// TIA Portal project "TrafficLight" (V19)

(* hardware
DEVICE "S7-1200 station_1"  S7-1200 Station
   slot 0: "Rack_0"  S7-1200 Rack  Rack  V1.0
   slot 1: "PLC_1"  CPU 1215C DC/DC/DC  6ES7 215-1AG40-0XB0  V4.6
*)

// ===== PLC "PLC_1"  CPU 1215C DC/DC/DC =====

VAR_GLOBAL   // PLC tag table "Default tag table"
   "emergencyButton" AT %I0.0 : Bool;
   "pedButtonDirB" AT %I0.1 : Bool;
   "pedButtonDirA" AT %I0.2 : Bool;
   "greenDirA" AT %Q0.0 : Bool;
   "yellowDirA" AT %Q0.1 : Bool;
   "redDirA" AT %Q0.2 : Bool;
   "pedGreenDirB" AT %Q0.3 : Bool;
   "pedRedDirB" AT %Q0.4 : Bool;
   "greenDirB" AT %Q0.5 : Bool;
   "yellowDirB" AT %Q0.6 : Bool;
   "redDirB" AT %Q0.7 : Bool;
   "pedGreenDirA" AT %Q1.0 : Bool;
   "pedRedDirA" AT %Q1.1 : Bool;
   "pedReqA" AT %M0.4 : Bool;
   "pedReqB" AT %M0.5 : Bool;
   "emergencyMode" AT %M0.6 : Bool;
   "current_dir" AT %M0.7 : Bool;
   "init_done" AT %M1.0 : Bool;
   "_debug" AT %M1.1 : Bool;
END_VAR

// folder: System blocks/Program resources

DATA_BLOCK "TP_Yellow_Phase_1"   // DB2
{ S7_Optimized_Access := 'TRUE' }
AUTHOR : Simatic
FAMILY : IEC
NAME : IEC_TMR
VERSION : 1.0
// stored: InstanceOfName IEC_TIMER
"IEC_TIMER"
BEGIN
END_DATA_BLOCK

DATA_BLOCK "TP_Yellow_Phase_2"   // DB3
{ S7_Optimized_Access := 'TRUE' }
AUTHOR : Simatic
FAMILY : IEC
NAME : IEC_TMR
VERSION : 1.0
// stored: InstanceOfName IEC_TIMER
"IEC_TIMER"
BEGIN
END_DATA_BLOCK

DATA_BLOCK "tp_main_loop"   // DB6
{ S7_Optimized_Access := 'TRUE' }
AUTHOR : Simatic
FAMILY : IEC
NAME : IEC_TMR
VERSION : 1.0
// stored: InstanceOfName IEC_TIMER
"IEC_TIMER"
BEGIN
END_DATA_BLOCK

DATA_BLOCK "ton_main_loop"   // DB7
{ S7_Optimized_Access := 'TRUE' }
AUTHOR : Simatic
FAMILY : IEC
NAME : IEC_TMR
VERSION : 1.0
// stored: InstanceOfName IEC_TIMER
"IEC_TIMER"
BEGIN
END_DATA_BLOCK

DATA_BLOCK "tp_main_loop_2"   // DB8
{ S7_Optimized_Access := 'TRUE' }
AUTHOR : Simatic
FAMILY : IEC
NAME : IEC_TMR
VERSION : 1.0
// stored: InstanceOfName IEC_TIMER
"IEC_TIMER"
BEGIN
END_DATA_BLOCK

// folder: (top level)

FUNCTION "ped_request" : Void   // FC1, LAD
{ S7_Optimized_Access := 'TRUE' }
VERSION : 0.1
   VAR_INPUT
      pred_A_or_B : String;
      ped_button : Bool;
      ped_req : Bool;
      ped_green : Bool;
      ped_red : Bool;
      dir_red : Bool;
   END_VAR
   VAR_OUTPUT
      o_ped_red : Bool;
      o_ped_green : Bool;
      o_ped_req : Bool;
   END_VAR
   VAR_TEMP
      r_trig_Q : Bool;
   END_VAR
   VAR_TEMP   // added for the SCL form of the ladder/FBD networks
      _w1 : Bool;
   END_VAR
BEGIN

REGION Network 1
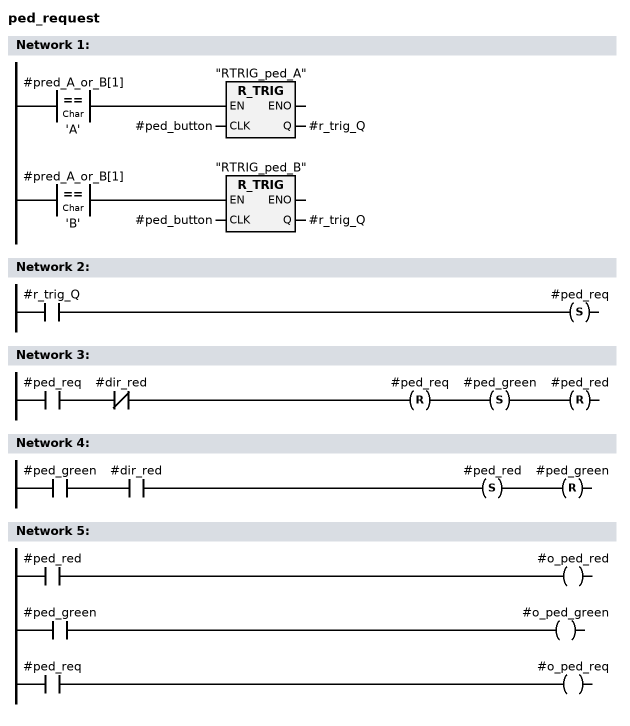
   IF #pred_A_or_B[1] = 'A' THEN
       "RTRIG_ped_A"(CLK := #ped_button, Q => #r_trig_Q);   // R_TRIG
   END_IF;
   IF #pred_A_or_B[1] = 'B' THEN
       "RTRIG_ped_B"(CLK := #ped_button, Q => #r_trig_Q);   // R_TRIG
   END_IF;
END_REGION

REGION Network 2
   RUNG wire#powerrail
      Contact( #r_trig_Q )
      S_Coil( #ped_req )
   END_RUNG
   // the same network as SCL:
   IF #r_trig_Q THEN #ped_req := TRUE; END_IF;
END_REGION

REGION Network 3
   RUNG wire#powerrail
      Contact( #ped_req )
      I_Contact( #dir_red )
      R_Coil( #ped_req )
      S_Coil( #ped_green )
      R_Coil( #ped_red )
   END_RUNG
   // the same network as SCL:
   #_w1 := #ped_req AND NOT #dir_red;
   IF #_w1 THEN
       #ped_req := FALSE;
       #ped_green := TRUE;
       #ped_red := FALSE;
   END_IF;
END_REGION

REGION Network 4
   RUNG wire#powerrail
      Contact( #ped_green )
      Contact( #dir_red )
      S_Coil( #ped_red )
      R_Coil( #ped_green )
   END_RUNG
   // the same network as SCL:
   IF #ped_green AND #dir_red THEN
       #ped_red := TRUE;
       #ped_green := FALSE;
   END_IF;
END_REGION

REGION Network 5
   RUNG wire#powerrail
      Contact( #ped_red )
      Coil( #o_ped_red )
   END_RUNG
   RUNG wire#powerrail
      Contact( #ped_green )
      Coil( #o_ped_green )
   END_RUNG
   RUNG wire#powerrail
      Contact( #ped_req )
      Coil( #o_ped_req )
   END_RUNG
   // the same network as SCL:
   #o_ped_red := #ped_red;
   #o_ped_green := #ped_green;
   #o_ped_req := #ped_req;
END_REGION
END_FUNCTION

FUNCTION "emerg" : Void   // FC2, LAD
{ S7_Optimized_Access := 'TRUE' }
VERSION : 0.1
   VAR_TEMP
      null_p : Bool;
   END_VAR
   VAR_TEMP   // added for the SCL form of the ladder/FBD networks
      _w1 : Bool;
      _w2 : Bool;
   END_VAR
BEGIN

REGION Network 1
   // Notice button click
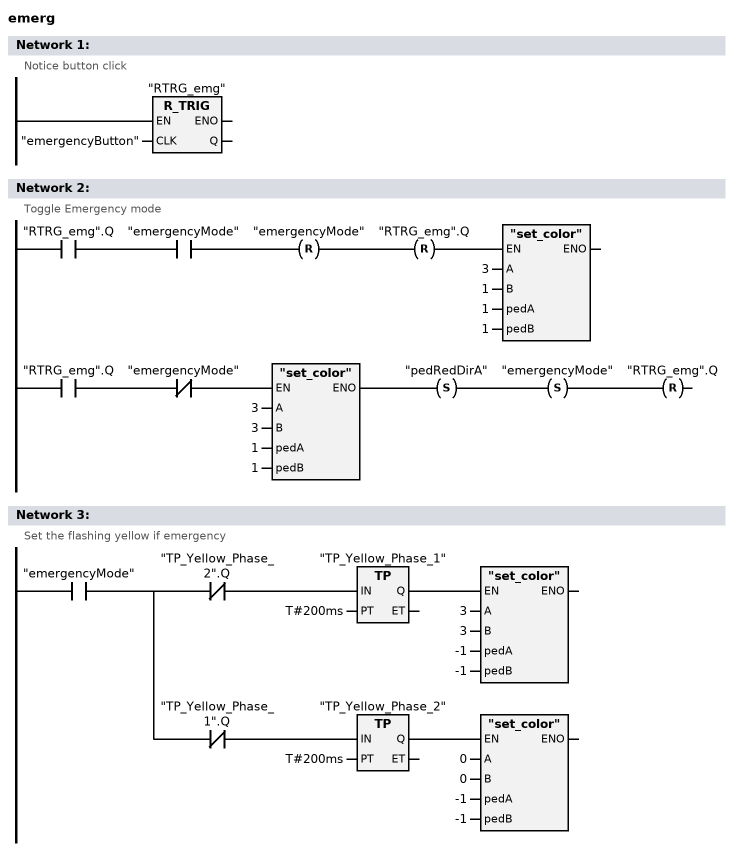
   "RTRG_emg"(CLK := "emergencyButton");   // R_TRIG
END_REGION

REGION Network 2
   // Toggle Emergency mode
   RUNG wire#powerrail
      Contact( "RTRG_emg".Q )
      Contact( "emergencyMode" )
      R_Coil( "emergencyMode" )
      R_Coil( "RTRG_emg".Q )
      "set_color"("A" := 3, "B" := 1, pedA := 1, pedB := 1)
   END_RUNG
   RUNG wire#powerrail
      Contact( "RTRG_emg".Q )
      I_Contact( "emergencyMode" )
      "set_color"("A" := 3, "B" := 3, pedA := 1, pedB := 1)
      S_Coil( "pedRedDirA" )
      S_Coil( "emergencyMode" )
      R_Coil( "RTRG_emg".Q )
   END_RUNG
   // the same network as SCL:
   #_w1 := "RTRG_emg".Q AND "emergencyMode";
   IF #_w1 THEN
       "emergencyMode" := FALSE;
       "RTRG_emg".Q := FALSE;
       "set_color"("A" := 3, "B" := 1, pedA := 1, pedB := 1);
   END_IF;
   "set_color"(EN := "RTRG_emg".Q AND NOT "emergencyMode",
               "A" := 3,
               "B" := 3,
               pedA := 1,
               pedB := 1,
               ENO => #_w2);
   IF #_w2 THEN
       "pedRedDirA" := TRUE;
       "emergencyMode" := TRUE;
       "RTRG_emg".Q := FALSE;
   END_IF;
END_REGION

REGION Network 3
   // Set the flashing yellow if emergency
   "TP_Yellow_Phase_1".TP(IN := "emergencyMode" AND NOT "TP_Yellow_Phase_2".Q, PT := T#200ms);
   #_w1 := "emergencyMode";
   IF "TP_Yellow_Phase_1".Q THEN "set_color"("A" := 3, "B" := 3, pedA := -1, pedB := -1); END_IF;
   "TP_Yellow_Phase_2".TP(IN := #_w1 AND NOT "TP_Yellow_Phase_1".Q, PT := T#200ms);
   IF "TP_Yellow_Phase_2".Q THEN "set_color"("A" := 0, "B" := 0, pedA := -1, pedB := -1); END_IF;
END_REGION
END_FUNCTION

FUNCTION "set_color" : Void   // FC3, LAD
{ S7_Optimized_Access := 'TRUE' }
VERSION : 0.1
// 1: red
// 2: green
// 3: yellow
// 
// 0: off
   VAR_INPUT
      "A" : Int;
      "B" : Int;
      pedA : Int;
      pedB : Int;
   END_VAR
BEGIN

REGION Network 1
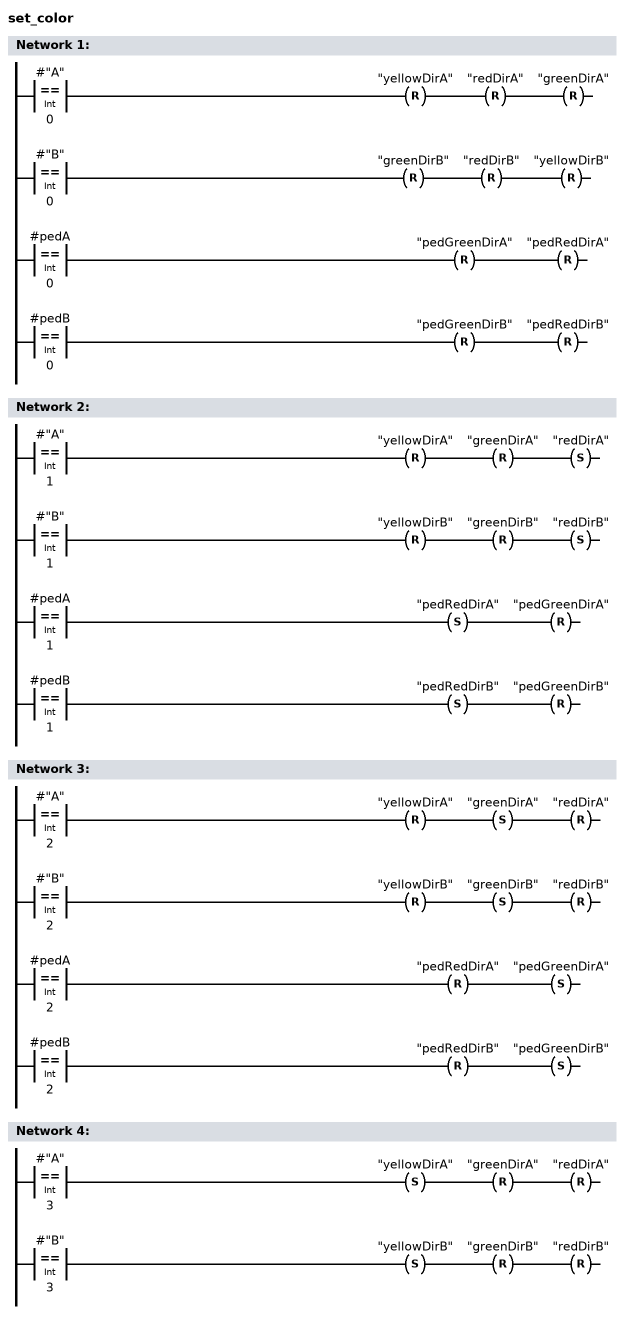
   RUNG wire#powerrail
      { S7_Templates := "SrcType := Int" } EQ_Contact(in1 := #"A", in2 := 0)
      R_Coil( "yellowDirA" )
      R_Coil( "redDirA" )
      R_Coil( "greenDirA" )
   END_RUNG
   RUNG wire#powerrail
      { S7_Templates := "SrcType := Int" } EQ_Contact(in1 := #"B", in2 := 0)
      R_Coil( "greenDirB" )
      R_Coil( "redDirB" )
      R_Coil( "yellowDirB" )
   END_RUNG
   RUNG wire#powerrail
      { S7_Templates := "SrcType := Int" } EQ_Contact(in1 := #pedA, in2 := 0)
      R_Coil( "pedGreenDirA" )
      R_Coil( "pedRedDirA" )
   END_RUNG
   RUNG wire#powerrail
      { S7_Templates := "SrcType := Int" } EQ_Contact(in1 := #pedB, in2 := 0)
      R_Coil( "pedGreenDirB" )
      R_Coil( "pedRedDirB" )
   END_RUNG
   // the same network as SCL:
   IF #"A" = 0 THEN
       "yellowDirA" := FALSE;
       "redDirA" := FALSE;
       "greenDirA" := FALSE;
   END_IF;
   IF #"B" = 0 THEN
       "greenDirB" := FALSE;
       "redDirB" := FALSE;
       "yellowDirB" := FALSE;
   END_IF;
   IF #pedA = 0 THEN
       "pedGreenDirA" := FALSE;
       "pedRedDirA" := FALSE;
   END_IF;
   IF #pedB = 0 THEN
       "pedGreenDirB" := FALSE;
       "pedRedDirB" := FALSE;
   END_IF;
END_REGION

REGION Network 2
   RUNG wire#powerrail
      { S7_Templates := "SrcType := Int" } EQ_Contact(in1 := #"A", in2 := 1)
      R_Coil( "yellowDirA" )
      R_Coil( "greenDirA" )
      S_Coil( "redDirA" )
   END_RUNG
   RUNG wire#powerrail
      { S7_Templates := "SrcType := Int" } EQ_Contact(in1 := #"B", in2 := 1)
      R_Coil( "yellowDirB" )
      R_Coil( "greenDirB" )
      S_Coil( "redDirB" )
   END_RUNG
   RUNG wire#powerrail
      { S7_Templates := "SrcType := Int" } EQ_Contact(in1 := #pedA, in2 := 1)
      S_Coil( "pedRedDirA" )
      R_Coil( "pedGreenDirA" )
   END_RUNG
   RUNG wire#powerrail
      { S7_Templates := "SrcType := Int" } EQ_Contact(in1 := #pedB, in2 := 1)
      S_Coil( "pedRedDirB" )
      R_Coil( "pedGreenDirB" )
   END_RUNG
   // the same network as SCL:
   IF #"A" = 1 THEN
       "yellowDirA" := FALSE;
       "greenDirA" := FALSE;
       "redDirA" := TRUE;
   END_IF;
   IF #"B" = 1 THEN
       "yellowDirB" := FALSE;
       "greenDirB" := FALSE;
       "redDirB" := TRUE;
   END_IF;
   IF #pedA = 1 THEN
       "pedRedDirA" := TRUE;
       "pedGreenDirA" := FALSE;
   END_IF;
   IF #pedB = 1 THEN
       "pedRedDirB" := TRUE;
       "pedGreenDirB" := FALSE;
   END_IF;
END_REGION

REGION Network 3
   RUNG wire#powerrail
      { S7_Templates := "SrcType := Int" } EQ_Contact(in1 := #"A", in2 := 2)
      R_Coil( "yellowDirA" )
      S_Coil( "greenDirA" )
      R_Coil( "redDirA" )
   END_RUNG
   RUNG wire#powerrail
      { S7_Templates := "SrcType := Int" } EQ_Contact(in1 := #"B", in2 := 2)
      R_Coil( "yellowDirB" )
      S_Coil( "greenDirB" )
      R_Coil( "redDirB" )
   END_RUNG
   RUNG wire#powerrail
      { S7_Templates := "SrcType := Int" } EQ_Contact(in1 := #pedA, in2 := 2)
      R_Coil( "pedRedDirA" )
      S_Coil( "pedGreenDirA" )
   END_RUNG
   RUNG wire#powerrail
      { S7_Templates := "SrcType := Int" } EQ_Contact(in1 := #pedB, in2 := 2)
      R_Coil( "pedRedDirB" )
      S_Coil( "pedGreenDirB" )
   END_RUNG
   // the same network as SCL:
   IF #"A" = 2 THEN
       "yellowDirA" := FALSE;
       "greenDirA" := TRUE;
       "redDirA" := FALSE;
   END_IF;
   IF #"B" = 2 THEN
       "yellowDirB" := FALSE;
       "greenDirB" := TRUE;
       "redDirB" := FALSE;
   END_IF;
   IF #pedA = 2 THEN
       "pedRedDirA" := FALSE;
       "pedGreenDirA" := TRUE;
   END_IF;
   IF #pedB = 2 THEN
       "pedRedDirB" := FALSE;
       "pedGreenDirB" := TRUE;
   END_IF;
END_REGION

REGION Network 4
   RUNG wire#powerrail
      { S7_Templates := "SrcType := Int" } EQ_Contact(in1 := #"A", in2 := 3)
      S_Coil( "yellowDirA" )
      R_Coil( "greenDirA" )
      R_Coil( "redDirA" )
   END_RUNG
   RUNG wire#powerrail
      { S7_Templates := "SrcType := Int" } EQ_Contact(in1 := #"B", in2 := 3)
      S_Coil( "yellowDirB" )
      R_Coil( "greenDirB" )
      R_Coil( "redDirB" )
   END_RUNG
   // the same network as SCL:
   IF #"A" = 3 THEN
       "yellowDirA" := TRUE;
       "greenDirA" := FALSE;
       "redDirA" := FALSE;
   END_IF;
   IF #"B" = 3 THEN
       "yellowDirB" := TRUE;
       "greenDirB" := FALSE;
       "redDirB" := FALSE;
   END_IF;
END_REGION
END_FUNCTION

FUNCTION "road_lights_loop" : Void   // FC4, LAD
{ S7_Optimized_Access := 'TRUE' }
VERSION : 0.1
   VAR_TEMP
      trans_p_green : Time;
      red_to_green_switch : Bool;
      yellow_to_red : Bool;
   END_VAR
   VAR CONSTANT
      phase_Green : Time := T#500MS;
      phase_Yellow : Time := T#200MS;
      phase_transition : Time := T#100MS;
   END_VAR
   VAR_TEMP   // added for the SCL form of the ladder/FBD networks
      _w1 : Bool;
      _w2 : Bool;
   END_VAR
BEGIN

REGION Network 1
   // all timers are off meaning start of round -> switch between dirs
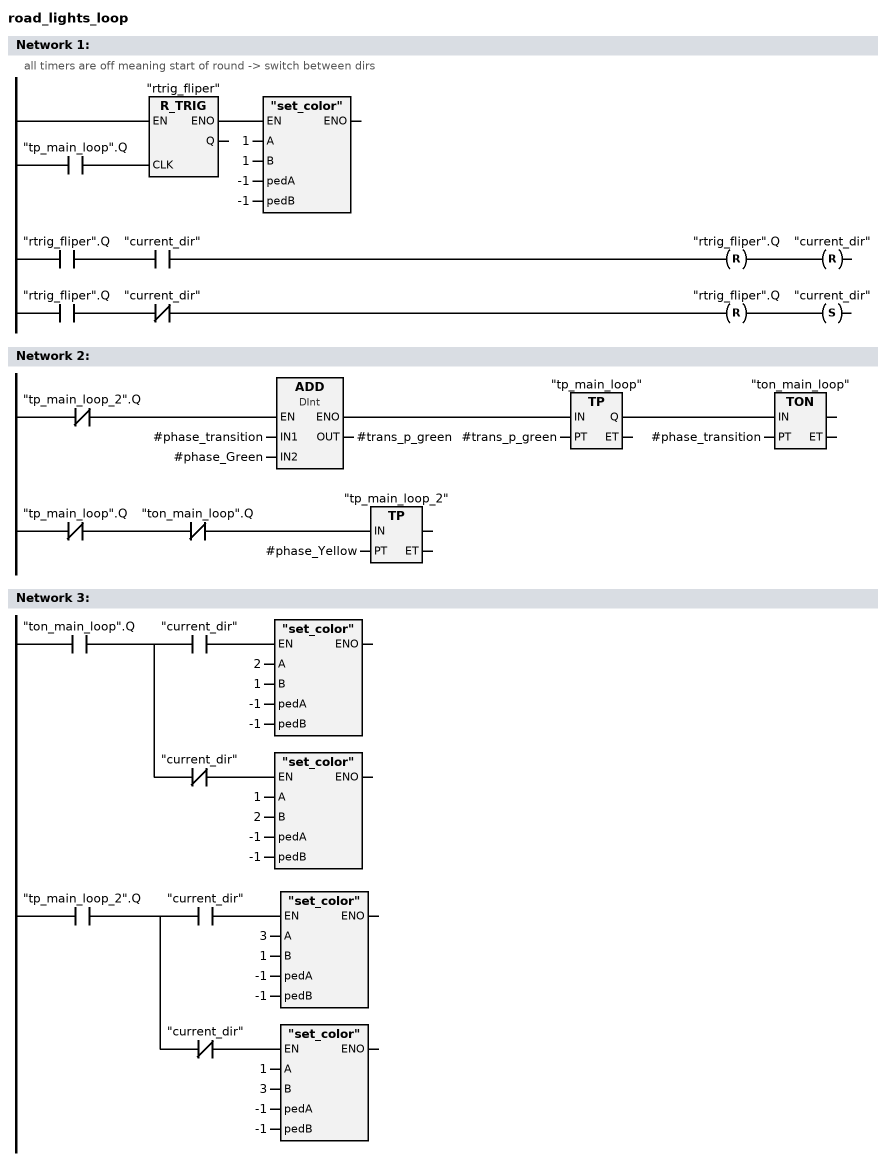
   // ENO of a box is taken as its EN; it also drops when the box reports an error
   "rtrig_fliper"(CLK := "tp_main_loop".Q);   // R_TRIG
   "set_color"("A" := 1, "B" := 1, pedA := -1, pedB := -1);
   #_w1 := "rtrig_fliper".Q AND "current_dir";
   IF #_w1 THEN
       "rtrig_fliper".Q := FALSE;
       "current_dir" := FALSE;
   END_IF;
   #_w2 := "rtrig_fliper".Q AND NOT "current_dir";
   IF #_w2 THEN
       "rtrig_fliper".Q := FALSE;
       "current_dir" := TRUE;
   END_IF;
END_REGION

REGION Network 2
   IF NOT "tp_main_loop_2".Q THEN #trans_p_green := #phase_transition + #phase_Green; END_IF;
   "tp_main_loop".TP(IN := NOT "tp_main_loop_2".Q, PT := #trans_p_green);
   "ton_main_loop".TON(IN := "tp_main_loop".Q, PT := #phase_transition);
   "tp_main_loop_2".TP(IN := NOT "tp_main_loop".Q AND NOT "ton_main_loop".Q, PT := #phase_Yellow);
END_REGION

REGION Network 3
   RUNG wire#powerrail
      Contact( "ton_main_loop".Q )
      wire#w1
      Contact( "current_dir" )
      "set_color"("A" := 2, "B" := 1, pedA := -1, pedB := -1)
   END_RUNG
   RUNG wire#w1
      I_Contact( "current_dir" )
      "set_color"("A" := 1, "B" := 2, pedA := -1, pedB := -1)
   END_RUNG
   RUNG wire#powerrail
      Contact( "tp_main_loop_2".Q )
      wire#w2
      Contact( "current_dir" )
      "set_color"("A" := 3, "B" := 1, pedA := -1, pedB := -1)
   END_RUNG
   RUNG wire#w2
      I_Contact( "current_dir" )
      "set_color"("A" := 1, "B" := 3, pedA := -1, pedB := -1)
   END_RUNG
   // the same network as SCL:
   #_w1 := "ton_main_loop".Q;
   IF "ton_main_loop".Q AND "current_dir" THEN
       "set_color"("A" := 2, "B" := 1, pedA := -1, pedB := -1);
   END_IF;
   IF #_w1 AND NOT "current_dir" THEN "set_color"("A" := 1, "B" := 2, pedA := -1, pedB := -1); END_IF;
   #_w2 := "tp_main_loop_2".Q;
   IF "tp_main_loop_2".Q AND "current_dir" THEN
       "set_color"("A" := 3, "B" := 1, pedA := -1, pedB := -1);
   END_IF;
   IF #_w2 AND NOT "current_dir" THEN "set_color"("A" := 1, "B" := 3, pedA := -1, pedB := -1); END_IF;
END_REGION
END_FUNCTION

ORGANIZATION_BLOCK "Main"   // OB1, LAD, ProgramCycle
TITLE = "Main Program Sweep (Cycle)"
{ S7_Optimized_Access := 'TRUE' }
VERSION : 0.1
   VAR_INPUT
      Initial_Call : Bool;   // Initial call of this OB
      Remanence : Bool;   // =True, if remanent data are available
   END_VAR
   VAR_TEMP   // added for the SCL form of the ladder/FBD networks
      _w1 : Bool;
   END_VAR
BEGIN

REGION Network 1
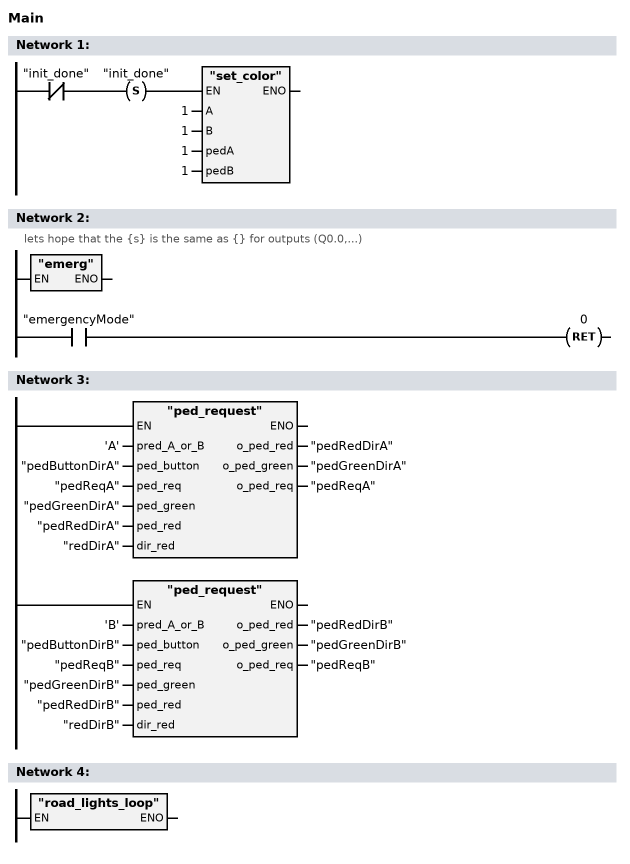
   RUNG wire#powerrail
      I_Contact( "init_done" )
      S_Coil( "init_done" )
      "set_color"("A" := 1, "B" := 1, pedA := 1, pedB := 1)
   END_RUNG
   // the same network as SCL:
   #_w1 := NOT "init_done";
   IF #_w1 THEN
       "init_done" := TRUE;
       "set_color"("A" := 1, "B" := 1, pedA := 1, pedB := 1);
   END_IF;
END_REGION

REGION Network 2
   // lets hope that the {s} is the same as {} for outputs (Q0.0,...)
   "emerg"();
   IF "emergencyMode" THEN
       ENO := 0;
       RETURN;
   END_IF;
END_REGION

REGION Network 3
   RUNG wire#powerrail
      "ped_request"(pred_A_or_B := 'A', ped_button := "pedButtonDirA", ped_req := "pedReqA", ped_green := "pedGreenDirA", ped_red := "pedRedDirA", dir_red := "redDirA", o_ped_red => "pedRedDirA", o_ped_green => "pedGreenDirA", o_ped_req => "pedReqA")
   END_RUNG
   RUNG wire#powerrail
      "ped_request"(pred_A_or_B := 'B', ped_button := "pedButtonDirB", ped_req := "pedReqB", ped_green := "pedGreenDirB", ped_red := "pedRedDirB", dir_red := "redDirB", o_ped_red => "pedRedDirB", o_ped_green => "pedGreenDirB", o_ped_req => "pedReqB")
   END_RUNG
   // the same network as SCL:
   "ped_request"(pred_A_or_B := 'A',
                 ped_button := "pedButtonDirA",
                 ped_req := "pedReqA",
                 ped_green := "pedGreenDirA",
                 ped_red := "pedRedDirA",
                 dir_red := "redDirA",
                 o_ped_red => "pedRedDirA",
                 o_ped_green => "pedGreenDirA",
                 o_ped_req => "pedReqA");
   "ped_request"(pred_A_or_B := 'B',
                 ped_button := "pedButtonDirB",
                 ped_req := "pedReqB",
                 ped_green := "pedGreenDirB",
                 ped_red := "pedRedDirB",
                 dir_red := "redDirB",
                 o_ped_red => "pedRedDirB",
                 o_ped_green => "pedGreenDirB",
                 o_ped_req => "pedReqB");
END_REGION

REGION Network 4
   RUNG wire#powerrail
      "road_lights_loop"()
   END_RUNG
   // the same network as SCL:
   "road_lights_loop"();
END_REGION
END_ORGANIZATION_BLOCK